SUBAPPLICATION Bool8_TO_logiBUS_QX8 (* 8 generische digitale Ausgaenge (Kanal frei waehlbar), gemeinsam getriggert durch 1 CNF-Event. Generisch fuer jede 8-Bit-Ausgangsgruppe. *)
  (* Standard: 61499-2 *)
  (* Version 1.0, 2026-09-09, Franz Höpfinger, Meisterschulen am Ostbahnhof, Ausgelagert aus Uebung_060_sub_Outputs (dort an TC-SC gebunden) - die 8 Ausgangskanaele waren zuvor fest importierte Output_Q1..Q8, jetzt als VarDeclaration parametrierbar zur Wiederverwendung fuer beliebige 8-Bit-Ausgangsgruppen. *)
  PACKAGE MyLib::sys;
  IMPORT logiBUS::io::DQ::logiBUS_DO;
  IMPORT logiBUS::io::DQ::logiBUS_DO_S;
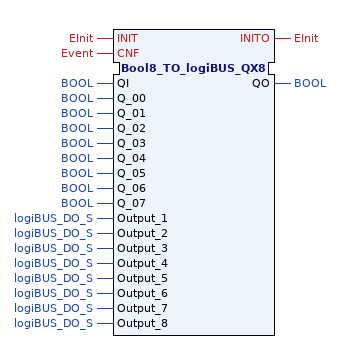
  EVENT_INPUT
    INIT : EInit; (* Initialization Request *)
    CNF;
  END_EVENT
  EVENT_OUTPUT
    INITO : EInit; (* Initialization Confirm *)
  END_EVENT
  VAR_INPUT
    QI : BOOL := TRUE; (* Quality Input - TRUE to enable service *)
    Q_00 : BOOL;
    Q_01 : BOOL;
    Q_02 : BOOL;
    Q_03 : BOOL;
    Q_04 : BOOL;
    Q_05 : BOOL;
    Q_06 : BOOL;
    Q_07 : BOOL;
    Output_1 : logiBUS::io::DQ::logiBUS_DO_S := logiBUS_DO::Invalid; (* Identify the Output Output_Q1..Q8 *)
    Output_2 : logiBUS::io::DQ::logiBUS_DO_S := logiBUS_DO::Invalid; (* Identify the Output Output_Q1..Q8 *)
    Output_3 : logiBUS::io::DQ::logiBUS_DO_S := logiBUS_DO::Invalid; (* Identify the Output Output_Q1..Q8 *)
    Output_4 : logiBUS::io::DQ::logiBUS_DO_S := logiBUS_DO::Invalid; (* Identify the Output Output_Q1..Q8 *)
    Output_5 : logiBUS::io::DQ::logiBUS_DO_S := logiBUS_DO::Invalid; (* Identify the Output Output_Q1..Q8 *)
    Output_6 : logiBUS::io::DQ::logiBUS_DO_S := logiBUS_DO::Invalid; (* Identify the Output Output_Q1..Q8 *)
    Output_7 : logiBUS::io::DQ::logiBUS_DO_S := logiBUS_DO::Invalid; (* Identify the Output Output_Q1..Q8 *)
    Output_8 : logiBUS::io::DQ::logiBUS_DO_S := logiBUS_DO::Invalid; (* Identify the Output Output_Q1..Q8 *)
  END_VAR
  VAR_OUTPUT
    QO : BOOL; (* Quality Output - TRUE if service executed successfully *)
  END_VAR
  FBS
    DigitalOutput_Q4 : logiBUS::io::DQ::logiBUS_QX;
    DigitalOutput_Q7 : logiBUS::io::DQ::logiBUS_QX;
    DigitalOutput_Q1 : logiBUS::io::DQ::logiBUS_QX;
    DigitalOutput_Q5 : logiBUS::io::DQ::logiBUS_QX;
    DigitalOutput_Q2 : logiBUS::io::DQ::logiBUS_QX;
    DigitalOutput_Q6 : logiBUS::io::DQ::logiBUS_QX;
    DigitalOutput_Q8 : logiBUS::io::DQ::logiBUS_QX;
    DigitalOutput_Q3 : logiBUS::io::DQ::logiBUS_QX;
    AND_QO : iec61131::booleanOperators::AND_BOOL_8;
  END_FBS
  EVENT_CONNECTIONS
    CNF TO DigitalOutput_Q4.REQ;
    CNF TO DigitalOutput_Q7.REQ;
    CNF TO DigitalOutput_Q1.REQ;
    CNF TO DigitalOutput_Q5.REQ;
    CNF TO DigitalOutput_Q2.REQ;
    CNF TO DigitalOutput_Q6.REQ;
    CNF TO DigitalOutput_Q8.REQ;
    CNF TO DigitalOutput_Q3.REQ;
    INIT TO DigitalOutput_Q4.INIT;
    DigitalOutput_Q4.INITO TO DigitalOutput_Q7.INIT;
    DigitalOutput_Q7.INITO TO DigitalOutput_Q1.INIT;
    DigitalOutput_Q1.INITO TO DigitalOutput_Q5.INIT;
    DigitalOutput_Q5.INITO TO DigitalOutput_Q2.INIT;
    DigitalOutput_Q2.INITO TO DigitalOutput_Q6.INIT;
    DigitalOutput_Q6.INITO TO DigitalOutput_Q8.INIT;
    DigitalOutput_Q8.INITO TO DigitalOutput_Q3.INIT;
    DigitalOutput_Q3.INITO TO INITO;
    DigitalOutput_Q3.INITO TO AND_QO.REQ;
  END_CONNECTIONS
  DATA_CONNECTIONS
    Q_06 TO DigitalOutput_Q7.OUT;
    Q_00 TO DigitalOutput_Q1.OUT;
    Q_04 TO DigitalOutput_Q5.OUT;
    Q_01 TO DigitalOutput_Q2.OUT;
    Q_05 TO DigitalOutput_Q6.OUT;
    Q_02 TO DigitalOutput_Q3.OUT;
    Q_03 TO DigitalOutput_Q4.OUT;
    Q_07 TO DigitalOutput_Q8.OUT;
    Output_1 TO DigitalOutput_Q1.Output;
    Output_2 TO DigitalOutput_Q2.Output;
    Output_3 TO DigitalOutput_Q3.Output;
    Output_4 TO DigitalOutput_Q4.Output;
    Output_5 TO DigitalOutput_Q5.Output;
    Output_6 TO DigitalOutput_Q6.Output;
    Output_7 TO DigitalOutput_Q7.Output;
    Output_8 TO DigitalOutput_Q8.Output;
    QI TO DigitalOutput_Q4.QI;
    QI TO DigitalOutput_Q7.QI;
    QI TO DigitalOutput_Q1.QI;
    QI TO DigitalOutput_Q5.QI;
    QI TO DigitalOutput_Q2.QI;
    QI TO DigitalOutput_Q6.QI;
    QI TO DigitalOutput_Q8.QI;
    QI TO DigitalOutput_Q3.QI;
    DigitalOutput_Q4.QO TO AND_QO.IN1;
    DigitalOutput_Q7.QO TO AND_QO.IN2;
    DigitalOutput_Q1.QO TO AND_QO.IN3;
    DigitalOutput_Q5.QO TO AND_QO.IN4;
    DigitalOutput_Q2.QO TO AND_QO.IN5;
    DigitalOutput_Q6.QO TO AND_QO.IN6;
    DigitalOutput_Q8.QO TO AND_QO.IN7;
    DigitalOutput_Q3.QO TO AND_QO.IN8;
    AND_QO.OUT TO QO;
  END_CONNECTIONS
END_SUBAPPLICATION
